FUNCTION_BLOCK SettleTime (* Basic Function Block Type *)
  (* Standard: 61499-2 *)
  (* Version 0.0, 10/6/2026, Schneider Electric, Template *)
  PACKAGE SE.Nereda;
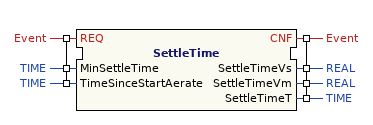
  EVENT_INPUT
    REQ WITH MinSettleTime, TimeSinceStartAerate; (* Normal Execution Request *)
  END_EVENT
  EVENT_OUTPUT
    CNF WITH SettleTimeVs, SettleTimeT, SettleTimeVm; (* Execution Confirmation *)
  END_EVENT
  VAR_INPUT
    MinSettleTime : TIME; (* Input event qualifier *)
    TimeSinceStartAerate : TIME;
  END_VAR
  VAR_OUTPUT
    SettleTimeVs : REAL; (* Output event qualifier *)
    SettleTimeVm : REAL;
    SettleTimeT : TIME;
  END_VAR
  VAR
    InMinSettleTime : REAL;
    InTimeSinceStartAerate : REAL;
    InSettleTimeV : REAL;
  END_VAR
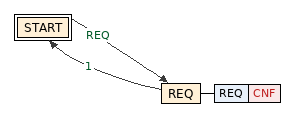
  EC_STATES
    START; (* Initial State *)
    REQ : REQ -> CNF; (* Normal execution *)
  END_STATES
  EC_TRANSITIONS
    START TO REQ := REQ;
    REQ TO START := 1;
  END_TRANSITIONS
  ALGORITHM REQ IN ST: (* Normally executed algorithm *)
;
InMinSettleTime := TIME_TO_REAL(MinSettleTime);
InTimeSinceStartAerate := TIME_TO_REAL(TimeSinceStartAerate);

InSettleTimeV := (InMinSettleTime - InTimeSinceStartAerate);

IF InSettleTimeV > 0 THEN
	SettleTimeVs := InSettleTimeV / 1000;
	SettleTimeT := REAL_TO_TIME(InSettleTimeV);
	SettleTimeVm := SettleTimeVs / 60;
ELSE
	SettleTimeVs := 0;
	SettleTimeVm := 0;
	SettleTimeT := T#0s;
END_IF;
  END_ALGORITHM
END_FUNCTION_BLOCK
